RoboDK station: Estacion_Final_TFG.rdk

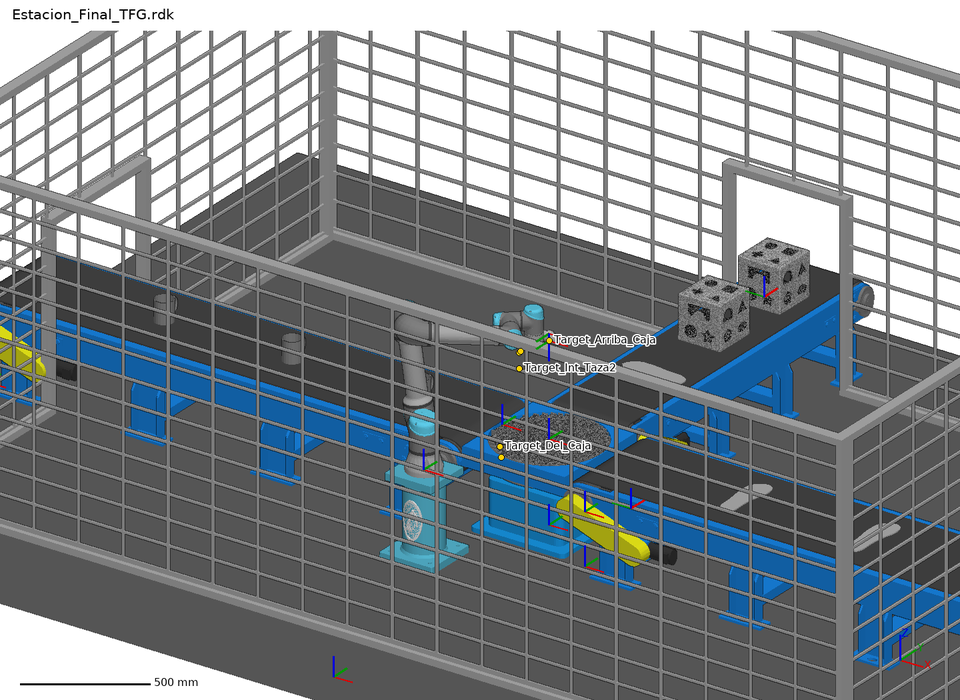
[picture v0: the station drawn from its stored meshes, robots at their saved joint values, targets as dots, program paths as lines]
Station Estacion_Final_TFG (saved by RoboDK 6.0.1). Poses are relative to the parent item; angles as X-Y-Z fixed-axis rotations.
Station parameters (name, value as stored): cara_actual, Cubo_Derecha, cam_delay, 0.005, contador, 10, prox_obj, Plantilla, defectuoso, 0, cont_def, 3, cont_ok, 4, prob_def, 5
  - folder Objetos
    - frame UR5e Base at (-167.75, -5.91, 0) mm
      - object Pedestal UR5 at (0, 0, -366.5) mm, size 250 x 250 x 366.5 mm, geometry from Pedestal-H12in-Type-1.sld
      - robot UR5e: 6 axes, payload 5 kg, reach 850 mm, repeatability 0.03 mm, weight 18.4 kg
          modified DH rows (alpha deg, a mm, theta deg, d mm): 0, 0, 0, 162.5; 90, 0, 180, 0; 0, 425, 0, 0; 0, 392.25, 0, 133.3; -90, 0, 0, 99.7; 90, 0, 180, 99.6
          joint limits [-360, -360, -360, -360, -360, -360] to [360, 360, 360, 360, 360, 360]; home [0, -90, -90, 0, 90, 0]; saved at [-138.346, -96.938, 101.969, -95.031, -90, -48.346]
        - frame Frame_Camara at (0, -105, 30.5) mm
          - camera Cámara 1
        - tool OnRobot Eyes Camera, TCP at (0.17, -105.19, 30.39) mm, size 104 x 155 x 41.9 mm
    - frame Frame_Cinta_Simple at (-2413.09, 275.71, -366.5) mm
      - robot Cinta_Simple: 1 axes
          modified DH rows (alpha deg, a mm, theta deg, d mm): 0, 0, 0, 0 linear
          base shift (0, 0, 0) mm, rotated rx 0 ry 90 rz 0 deg
          joint limits [-900000] to [900000]; home [0]; saved at [6082.39]
        - frame Frame_Padre_Cinta at (-2.39, 215, 0) mm
          - object Taza8 at (-4200, 0, 0) mm, rotated rx 0 ry 0 rz 90 deg, size 123.1 x 83.9 x 97 mm, geometry from Taza_Base.stp
          - object Taza9 at (-4800, 0, 0) mm, rotated rx 0 ry 0 rz 90 deg, size 123.1 x 83.9 x 97 mm, geometry from Taza_Base.stp
          - object Taza10 at (-5400, 0, 0) mm, rotated rx 0 ry 0 rz 90 deg, size 123.1 x 83.9 x 97 mm, geometry from Taza_Base.stp
    - frame Frame_Obj_Ref at (0, -850, -500) mm
      - object Juguete_ni at (0, 0, 0) mm, size 200 x 200 x 200 mm, geometry from Juguete_niños.stp
      - object Juguete_ni at (0, 0, 0) mm, size 200 x 200 x 200 mm, geometry from Juguete_niños_Arriba.stp
      - object Juguete_ni at (0, 0, 0) mm, size 200 x 200 x 200 mm, geometry from Juguete_niños_Der.stp
      - object Juguete_ni at (0, 0, 0) mm, size 200 x 200 x 200 mm, geometry from Juguete_niños_Frente.stp
      - object Juguete_ni at (0, 0, 0) mm, size 200 x 200 x 200 mm, geometry from Juguete_niños_Izq.stp
      - object Juguete_ni at (0, 0, 0) mm, size 200 x 200 x 200 mm, geometry from Juguete_niños_Det.stp
      - object Taza_Base at (0, 0, 0) mm, rotated rx 0 ry 0 rz 90 deg, size 123.1 x 83.9 x 97 mm, geometry from Taza_Base.stp
      - object Taza_Def1 at (0, 0, 0) mm, rotated rx 0 ry 0 rz 90 deg, size 123.1 x 83.9 x 97 mm, geometry from Taza_DibujoMal.stp
      - object Taza_Def2 at (0, 0, 0) mm, rotated rx 0 ry 0 rz 90 deg, size 123.1 x 83.9 x 97 mm, geometry from Taza_FaltaLetra.stp
      - object Plantilla_Derecha_Bien at (0, 0, 0) mm, rotated rx 90 ry 0 rz 0 deg, size 99.5 x 5 x 284.6 mm, geometry from Plantilla_Derecha_Bien.stl
      - object Plantilla_Derecha_Def1 at (0, 0, 0) mm, rotated rx 90 ry 0 rz 0 deg, size 99.6 x 5 x 284.5 mm, geometry from Plantilla_Derecha_Mal_Corte_Arriba.stl
      - object Plantilla_Derecha_Def2 at (0, 0, 0) mm, rotated rx 90 ry 0 rz 0 deg, size 99.6 x 5 x 284.6 mm, geometry from Plantilla_Derecha_Mal_Muescas.stl
      - object Plantilla_Izquierda_Bien at (0, 0, 0) mm, rotated rx 90 ry 0 rz 0 deg, size 99.5 x 5 x 284.6 mm, geometry from Plantilla_Izquierda_Bien.stl
      - object Plantilla_Izquierda_Def1 at (0, 0, 0) mm, rotated rx 90 ry 0 rz 0 deg, size 99.5 x 5 x 283.3 mm, geometry from Plantilla_Izquierda_Mal_Corte_Abajo.stl
      - object Plantilla_Izquierda_Def2 at (0, 0, 0) mm, rotated rx 90 ry 0 rz 0 deg, size 99.6 x 5 x 284.6 mm, geometry from Plantilla_Izquierda_Mal_Muescas.stl
    - frame Mesa_Rotatoria Base at (71.91, 490.71, -366.5) mm
      - robot Mesa_Rotatoria: 1 axes
          modified DH rows (alpha deg, a mm, theta deg, d mm): 0, 0, 0, 0
          joint limits [-360] to [360]; home [0]; saved at [0]
        - frame Cinta_Rotativa Base at (-220, 0, 366.5) mm
          - robot Cinta_Rotativa: 1 axes
              modified DH rows (alpha deg, a mm, theta deg, d mm): 0, 0, 0, 0 linear
              base shift (0, 0, 0) mm, rotated rx 0 ry 90 rz 0 deg
              joint limits [-10000] to [10000]; home [0]; saved at [3080]
      - object Base_Cinta at (0, 0, 280) mm, size 480 x 480 x 86.5 mm, geometry from Base_Cinta.stp
    - frame Frame_Cinta_OK at (391.91, 270.71, -366.5) mm
      - robot Cinta_OK: 1 axes
          modified DH rows (alpha deg, a mm, theta deg, d mm): 0, 0, 0, 0 linear
          base shift (0, 0, 0) mm, rotated rx 0 ry 90 rz 0 deg
          joint limits [-900000] to [900000]; home [0]; saved at [2400]
        - frame Frame_Padre_Cinta_OK at (-2.39, 215, 0) mm
          - object OK2 at (-600, 0, 0) mm, size 200 x 200 x 200 mm, geometry from Juguete_niños.stp
          - object OK3 at (-1200, 0, 0) mm, rotated rx 90 ry 0 rz 0 deg, size 99.5 x 5 x 284.6 mm, geometry from Plantilla_Izquierda_Bien.stl
          - object OK4 at (-1800, 0, 0) mm, rotated rx 90 ry 0 rz 0 deg, size 99.5 x 5 x 284.6 mm, geometry from Plantilla_Izquierda_Bien.stl
    - frame Frame_Cinta_Def at (247.91, 787.71, -366.5) mm, rotated rx 0 ry 0 rz 90 deg
      - robot Cinta_Def: 1 axes
          modified DH rows (alpha deg, a mm, theta deg, d mm): 0, 0, 0, 0 linear
          base shift (0, 0, 0) mm, rotated rx 0 ry 90 rz 0 deg
          joint limits [-900000] to [900000]; home [0]; saved at [1200]
        - frame Frame_Padre_Cinta_Def at (-2.39, 215, 0) mm
          - object Defectuoso1 at (0, -44, 0) mm, size 200 x 200 x 200 mm, geometry from Juguete_niños_Det.stp
          - object Defectuoso2 at (-400, -44, 0) mm, size 200 x 200 x 200 mm, geometry from Juguete_niños_Det.stp
          - object Defectuoso3 at (-800, -44, 0) mm, rotated rx 90 ry 0 rz 0 deg, size 99.6 x 5 x 284.5 mm, geometry from Plantilla_Derecha_Mal_Corte_Arriba.stl
    - frame Frame_Suelo at (117.25, 664.09, -367) mm
      - object Suelo at (0, 0, 0) mm, size 5420 x 3890 x 0 mm, geometry from Floor.sld
  - frame Frame_Targets at (71.91, 490.71, 450) mm, rotated rx 180 ry 0 rz 0 deg
    - target Target_Arriba_Caja (Cartesian target) at (0, 0, 30) mm; joints [-138.346, -96.938, 101.969, -95.031, -90, -48.346] of UR5e
    - target Target_Del_Caja (Cartesian target) at (0, 330, 350) mm, rotated rx 90 ry 0 rz 0 deg; joints [-204.685, -47.932, 150.066, -102.134, -24.685, -180] of UR5e
    - target Target_Int_Del (Cartesian target) at (0, 200, 0) mm; joints [-168.17, -117.089, 115.815, -88.726, -90, -78.17] of UR5e
    - target Target_Int_Taza1 (Cartesian target) at (0, 190, 0) mm; joints [-165.144, -119.371, 116.87, -87.498, -90, -75.144] of UR5e
    - target Target_Int_Taza2 (Cartesian target) at (0, 200, 70) mm, rotated rx 60 ry 0 rz 0 deg; joints [-180.443, -119.916, 146.516, -115.834, -30.003, -90.885] of UR5e
    - target Target_Taza (Cartesian target) at (0, 320, 400) mm, rotated rx 90 ry 0 rz 0 deg; joints [-202.098, -35.728, 146.743, -111.015, -22.098, -180] of UR5e
  - frame Frame_Target_Mesa at (71.91, 490.71, 0) mm
    - target Init_Mesa (Cartesian target) at (0, 0, 0) mm; joints [0, -47.932, 150.066, -102.134, -24.685, -180] of Mesa_Rotatoria
    - target Cubo_Izq (Cartesian target) at (0, 0, 0) mm, rotated rx 0 ry 0 rz 90 deg; joints [90, -47.932, 150.066, -102.134, -24.685, -180] of Mesa_Rotatoria
    - target Cubo_Detras (Cartesian target) at (0, 0, 0) mm, rotated rx 0 ry 0 rz 180 deg; joints [180, -47.932, 150.066, -102.134, -24.685, -180] of Mesa_Rotatoria
    - target Cubo_Der (Cartesian target) at (0, 0, 0) mm, rotated rx 0 ry 0 rz -90 deg; joints [270, -47.932, 150.066, -102.134, -24.685, -180] of Mesa_Rotatoria
    - target Target_Def (Cartesian target) at (0, 0, 0) mm, rotated rx 0 ry 0 rz 90 deg; joints [90, -47.932, 150.066, -102.134, -24.685, -180] of Mesa_Rotatoria
    - target Target_Taza_Mesa (Cartesian target) at (0, 0, 0) mm, rotated rx 0 ry 0 rz 90 deg; joints [90, -47.932, 150.066, -102.134, -24.685, -180] of Mesa_Rotatoria
  - folder Vallado
    - frame Frame Valla Trasera at (2332.25, -755.91, -366.5) mm, rotated rx 0 ry 0 rz 90 deg
      - object VallaTrasera at (0, 0, 0) mm, rotated rx 90 ry 0 rz 90 deg, size 4420 x 1500 x 50 mm, geometry from VallaBigCap.stl
    - frame Frame Valla Entrada at (-2062.75, -730.91, -366.5) mm, rotated rx 0 ry 0 rz -90 deg
      - object Valla_Entrada at (0, 0, 0) mm, rotated rx 90 ry 0 rz 180 deg, size 2790 x 1500 x 50 mm, geometry from Valla_Enrada.stp
    - frame Frame Valla Salida at (2307.25, -730.91, -366.5) mm, rotated rx 0 ry 0 rz -90 deg
      - object Valla_Salida at (0, 0, 0) mm, rotated rx 90 ry 0 rz 180 deg, size 2790 x 1500 x 50 mm, geometry from Valla_Enrada.stp
    - frame Frame Valla Defectuosas at (2332.25, 2084.09, -366.5) mm, rotated rx 0 ry 0 rz 180 deg
      - object Valla_CintaDef at (0, 0, 0) mm, rotated rx 90 ry 0 rz 0 deg, size 4420 x 1500 x 50 mm, geometry from Valla_CintaDef.stp
  - folder Programas
    - Python program Global (listed below)
    - Python program Reset (listed below)
  - folder Comparacion
    - Python program Comp_Inicial (listed below)
    - Python program Comp_Plantilla (listed below)
    - folder Codigos Cubo
      - Python program Comp_Cubo (listed below)
      - Python program Cubo_General (listed below)
    - folder Codigos Taza
      - Python program Comp_Taza (listed below)
      - Python program Taza_General (listed below)
  - folder Cintas
    - Python program Generar_Objeto (listed below)
    - Python program Avanzar_Cinta_Rot (listed below)

--- Python program Global ---
# Type help("robodk.robolink") or help("robodk.robomath") for more information
# Press F5 to run the script
# Documentation: https://robodk.com/doc/en/RoboDK-API.html
# Reference:     https://robodk.com/doc/en/PythonAPI/robodk.html
# Note: It is not required to keep a copy of this file, your Python script is saved with your RDK project

# You can also use the new version of the API:
from robodk import *      # RoboDK API
from robolink import *    # Robot toolbox
RDK = robolink.Robolink()

robot = RDK.Item('UR5e')
tool = RDK.Item('OnRobot Eyes Camera')
frame_target = RDK.Item('Frame_Targets')
init = RDK.Item('Reset')
avanzarCinta = RDK.Item('Generar_Objeto')
frame_mesa = RDK.Item('Frame_Target_Mesa')

arriba = RDK.Item('Target_Arriba_Caja')

robot.setPoseFrame(frame_target)
robot.MoveJ(arriba)

mesa=RDK.Item('Mesa_Rotatoria',itemtype=ITEM_TYPE_ROBOT)
cinta_rot=RDK.Item('Cinta_Rotativa',itemtype=ITEM_TYPE_ROBOT)
cinta_ok=RDK.Item('Cinta_OK',itemtype=ITEM_TYPE_ROBOT)
cinta_def=RDK.Item('Cinta_Def',itemtype=ITEM_TYPE_ROBOT)
ident = RDK.Item('Comp_Inicial')
comp_plantilla = RDK.Item('Comp_Plantilla')
comp_cubo = RDK.Item('Cubo_General')
comp_taza = RDK.Item('Taza_General')
avanzar_cinta_rot = RDK.Item('Avanzar_Cinta_Rot')
init_mesa = RDK.Item('Init_Mesa')
pos_def = RDK.Item('Target_Def')


frame_padre_def=RDK.Item('Frame_Padre_Cinta_Def')
frame_padre_ok=RDK.Item('Frame_Padre_Cinta_OK')

mesa.setPoseFrame(frame_mesa)

init.RunProgram()
init.WaitFinished()
obj_scan = RDK.getParam('prox_obj')

while True:
    while obj_scan == 'NULL':
        avanzarCinta.RunProgram()
        avanzarCinta.WaitFinished()
        obj_scan = RDK.getParam('prox_obj')

    avanzar_cinta_rot.RunProgram()
    avanzar_cinta_rot.WaitFinished()

    ident.RunProgram()
    ident.WaitFinished()

    defecto = RDK.getParam('defectuoso')
    contador = int(RDK.getParam('contador'))
    contador_def = int(RDK.getParam('cont_def'))
    contador_ok = int(RDK.getParam('cont_ok'))
    nombre_obj = obj_scan+str(contador-3)
    obj_listo = RDK.Item(nombre_obj)

    if defecto == 1:
        mesa.MoveJ(pos_def)
        avanzar_cinta_rot.RunProgram()
        avanzar_cinta_rot.WaitFinished()
        obj_listo.setParent(frame_padre_def)
        if obj_scan == 'Plantilla':
            obj_listo.setPose(transl((-400*(contador_def)),-44,0) * rotx(pi/2))
        elif obj_scan == 'Taza':
            obj_listo.setPose(transl((-400*(contador_def)),-44,0) * rotz(pi/2))
        else:
            obj_listo.setPose(transl((-400*(contador_def)),-44,0))
        cinta_def.MoveJ(cinta_def.Joints()+400)
        contador_def += 1
        obj_listo.setName('Defectuoso'+str(contador_def))
        if contador_def > 3:
            obj_borrar = RDK.Item('Defectuoso'+str(contador_def-3))
            RDK.Delete(obj_borrar)

    else:
        mesa.MoveJ(init_mesa)
        avanzar_cinta_rot.RunProgram()
        avanzar_cinta_rot.WaitFinished()
        obj_listo.setParent(frame_padre_ok)
        if obj_scan == 'Plantilla':
            obj_listo.setPose(transl((-600*(contador_ok)),0,0) * rotx(pi/2))
        elif obj_scan == 'Taza':
            obj_listo.setPose(transl((-600*(contador_ok)),0,0) * rotz(pi/2))
        else:
            obj_listo.setPose(transl((-600*(contador_ok)),0,0))
        cinta_ok.MoveJ(cinta_ok.Joints()+600)
        contador_ok += 1
        obj_listo.setName('OK'+str(contador_ok))
        if contador_ok > 3:
            obj_borrar = RDK.Item('OK'+str(contador_ok-3))
            RDK.Delete(obj_borrar)

    RDK.setParam('cont_def',contador_def)
    RDK.setParam('cont_ok',contador_ok)
    mesa.MoveJ(init_mesa)
    RDK.setParam('defectuoso',0)
    avanzarCinta.RunProgram()
    avanzarCinta.WaitFinished()
    obj_scan = RDK.getParam('prox_obj')

--- Python program Reset ---
# Type help("robodk.robolink") or help("robodk.robomath") for more information
# Press F5 to run the script
# Documentation: https://robodk.com/doc/en/RoboDK-API.html
# Reference:     https://robodk.com/doc/en/PythonAPI/robodk.html
# Note: It is not required to keep a copy of this file, your Python script is saved with your RDK project

import random

# Forward and backwards compatible use of the RoboDK API:
# Remove these 2 lines to follow python programming guidelines
from robodk import *      # RoboDK API
from robolink import *    # Robot toolbox
# Link to RoboDK
RDK = Robolink()

num=random.randint(1,3)
#num=3

RDK.setParam('contador',1)
RDK.setParam('cont_def',0)
RDK.setParam('cont_ok',0)
RDK.setParam('defectuoso',0)

if num == 1: # Caso de que sea plantilla
    num2 = random.randint(1,2)
    if num2 == 1: # Plantilla izquierda
        num3 = random.randint(1,6)
        if num3 == 5: # Defecto 1
            padre = RDK.Item('Plantilla_Izquierda_Def1')
            nombreCopia = 'Plantilla'
        elif num3 == 6: # Defecto 2
            padre = RDK.Item('Plantilla_Izquierda_Def2')
            nombreCopia = 'Plantilla'
        else:
            padre = RDK.Item('Plantilla_Izquierda_Bien')
            nombreCopia = 'Plantilla'
    if num2 == 2: # Plantilla izquierda
        num3 = random.randint(1,6)
        if num3 == 5: # Defecto 1
            padre = RDK.Item('Plantilla_Derecha_Def1')
            nombreCopia = 'Plantilla'
        elif num3 == 6: # Defecto 2
            padre = RDK.Item('Plantilla_Derecha_Def2')
            nombreCopia = 'Plantilla'
        else:
            padre = RDK.Item('Plantilla_Derecha_Bien')
            nombreCopia = 'Plantilla'

elif num == 2: # Caso de que sea Juguete
    num2 = random.randint(1,10)
    if num2 == 6: # Juguete mal arriba
        padre = RDK.Item('Juguete_niños_Arriba')
        nombreCopia = 'Juguete_niños'
    elif num2 == 7: # Juguete mal izquierda
        padre = RDK.Item('Juguete_niños_Izq')
        nombreCopia = 'Juguete_niños'
    elif num2 == 8: # Juguete mal derecha
        padre = RDK.Item('Juguete_niños_Der')
        nombreCopia = 'Juguete_niños'
    elif num2 == 9: # Juguete mal delante
        padre = RDK.Item('Juguete_niños_Del')
        nombreCopia = 'Juguete_niños'
    elif num2 == 10: # Juguete mal detras
        padre = RDK.Item('Juguete_niños_Det')
        nombreCopia = 'Juguete_niños'
    else: # Caso sin fallos
        padre = RDK.Item('Juguete_niños_Base')
        nombreCopia = 'Juguete_niños'

elif num == 3: # Caso de que sea taza
    num2 = random.randint(1,6)
    if num2 == 5: # Defecto 1
        padre = RDK.Item('Taza_Def1')
        nombreCopia = 'Taza'
    elif num2 == 6: # Defecto 2
        padre = RDK.Item('Taza_Def2')
        nombreCopia = 'Taza'
    else:
        padre = RDK.Item('Taza_Base')
        nombreCopia = 'Taza'


MECHANISM_NAME = 'Cinta_Simple'
mechanism=RDK.Item(MECHANISM_NAME,itemtype=ITEM_TYPE_ROBOT)
cinta_ok=RDK.Item('Cinta_OK',itemtype=ITEM_TYPE_ROBOT)
cinta_def=RDK.Item('Cinta_Def',itemtype=ITEM_TYPE_ROBOT)
cinta_rot=RDK.Item('Cinta_Rotativa',itemtype=ITEM_TYPE_ROBOT)
frame_padre_def=RDK.Item('Frame_Padre_Cinta_Def')
frame_padre_ok=RDK.Item('Frame_Padre_Cinta_OK')
mesa = RDK.Item('Mesa_Rotatoria')

frame_padre=RDK.Item('Frame_Padre_Cinta')

if mechanism.Valid() and cinta_rot.Valid() and mesa.Valid():
    mechanism.setJoints([467.39])
    cinta_ok.setJoints([0])
    cinta_def.setJoints([0])
    cinta_rot.setJoints([0])
    mesa.setJoints([0])
    RDK.Delete(frame_padre.Childs())
    RDK.Delete(frame_padre_def.Childs())
    RDK.Delete(frame_padre_ok.Childs())
    RDK.Delete(cinta_rot.Childs())
    padre.Copy()
    copia=RDK.Paste()
    copia.setParent(frame_padre)
    RDK.setParam('prox_obj','NULL')
    #hacemos visible el objeto nuevo
    cont = int(RDK.getParam('contador'))
    copia.setName(nombreCopia+str(cont))
    copia.setVisible(1)

--- Python program Comp_Inicial ---
from robolink import *
import cv2 as cv
import numpy as np
import os

RDK = Robolink()
cam_item = RDK.Item('Cámara 1', ITEM_TYPE_CAMERA)
carpeta = r"C:\Users\algob\OneDrive\UPV\4 - Cuarto\TFG\Imagen"

comp_plantilla = RDK.Item('Comp_Plantilla')
comp_cubo = RDK.Item('Cubo_General')
comp_taza = RDK.Item('Taza_General')

# 1. Cargar las dos imagenes de referencia en escala de grises (RAW)
img_izq_raw = cv.imread(os.path.join(carpeta, "Ref_izq.png"), 0)
img_der_raw = cv.imread(os.path.join(carpeta, "Ref_der.png"), 0)
img_cubo_raw = cv.imread(os.path.join(carpeta, "Cubo", "Cubo_Arriba_base.png"), 0)
img_taza_raw = cv.imread(os.path.join(carpeta, "Taza", "Taza_Arriba.png"), 0)

# FILTRO: Convertir el fondo gris en NEGRO puro y la plantilla en BLANCO puro
_, img_izq = cv.threshold(img_izq_raw, 200, 255, cv.THRESH_BINARY)
_, img_der = cv.threshold(img_der_raw, 200, 255, cv.THRESH_BINARY)
_, img_cubo = cv.threshold(img_cubo_raw, 200, 255, cv.THRESH_BINARY)
_, img_taza = cv.threshold(img_taza_raw, 200, 255, cv.THRESH_BINARY)

def obtener_contorno_principal(img_bw):
    # RETR_EXTERNAL busca únicamente el contorno exterior más externo
    cnts, _ = cv.findContours(img_bw, cv.RETR_EXTERNAL, cv.CHAIN_APPROX_SIMPLE)
    return max(cnts, key=cv.contourArea) if cnts else None

ref_izq = obtener_contorno_principal(img_izq)
ref_der = obtener_contorno_principal(img_der)
ref_cubo = obtener_contorno_principal(img_cubo)
ref_taza = obtener_contorno_principal(img_taza)

tiempo_inicio = time.time()
DURACION_MAXIMA = RDK.getParam('cam_delay')

while True:
    if (time.time() - tiempo_inicio) > DURACION_MAXIMA:
        cv.destroyAllWindows()
        cv.waitKey(1)
        break

    bytes_img = RDK.Cam2D_Snapshot("", cam_item)
    if bytes_img == b'':
        cv.destroyAllWindows()
        cv.waitKey(1)
        break

    img = cv.imdecode(np.frombuffer(bytes_img, np.uint8), cv.IMREAD_UNCHANGED)
    gray = cv.cvtColor(img, cv.COLOR_BGR2GRAY)

    _, thresh = cv.threshold(gray, 200, 255, cv.THRESH_BINARY)
    actual = obtener_contorno_principal(thresh)

    if actual is not None:
        diff_izq = cv.matchShapes(ref_izq, actual, 1, 0.0)
        diff_der = cv.matchShapes(ref_der, actual, 1, 0.0)
        diff_cubo = cv.matchShapes(ref_cubo, actual, 1, 0.0)
        diff_taza = cv.matchShapes(ref_taza, actual, 1, 0.0)

        mejor_diff = min(diff_izq, diff_der, diff_taza, diff_cubo)

        if mejor_diff == diff_izq or mejor_diff == diff_der:
            comp_plantilla.RunProgram()
            comp_plantilla.WaitFinished()
        elif mejor_diff == diff_cubo:
            comp_cubo.RunProgram()
            comp_cubo.WaitFinished()
        elif mejor_diff == diff_taza:
            comp_taza.RunProgram()
            comp_taza.WaitFinished()

cv.destroyAllWindows()
cv.waitKey(1)

--- Python program Comp_Plantilla ---
from robolink import *
import cv2 as cv
import numpy as np
import os

RDK = Robolink()
cam_item = RDK.Item('Cámara 1', ITEM_TYPE_CAMERA)
carpeta = r"C:\Users\algob\OneDrive\UPV\4 - Cuarto\TFG\Imagen"

# 1. Cargar las dos imagenes de referencia en escala de grises (RAW)
img_izq_raw = cv.imread(os.path.join(carpeta, "Ref_izq.png"), 0)
img_der_raw = cv.imread(os.path.join(carpeta, "Ref_der.png"), 0)

# FILTRO: Convertir el fondo gris en NEGRO puro y la plantilla en BLANCO puro
_, img_izq = cv.threshold(img_izq_raw, 200, 255, cv.THRESH_BINARY)
_, img_der = cv.threshold(img_der_raw, 200, 255, cv.THRESH_BINARY)

def obtener_contorno_principal(img_bw):
    # RETR_EXTERNAL busca únicamente el contorno exterior más externo
    cnts, _ = cv.findContours(img_bw, cv.RETR_EXTERNAL, cv.CHAIN_APPROX_SIMPLE)
    return max(cnts, key=cv.contourArea) if cnts else None

ref_izq = obtener_contorno_principal(img_izq)
ref_der = obtener_contorno_principal(img_der)

# Umbral de aceptación
UMBRAL = 0.01
tiempo_inicio = time.time()
DURACION_MAXIMA = RDK.getParam('cam_delay')

while True:
    if (time.time() - tiempo_inicio) > DURACION_MAXIMA:
        cv.destroyAllWindows()
        cv.waitKey(1)
        break

    bytes_img = RDK.Cam2D_Snapshot("", cam_item)
    if bytes_img == b'':
        cv.destroyAllWindows()
        cv.waitKey(1)
        break

    img = cv.imdecode(np.frombuffer(bytes_img, np.uint8), cv.IMREAD_UNCHANGED)
    gray = cv.cvtColor(img, cv.COLOR_BGR2GRAY)

    _, thresh = cv.threshold(gray, 200, 255, cv.THRESH_BINARY)
    actual = obtener_contorno_principal(thresh)

    if actual is not None:
        # 2. Comparar con ambas imagenes de referencia
        diff_izq = cv.matchShapes(ref_izq, actual, 1, 0.0)
        diff_der = cv.matchShapes(ref_der, actual, 1, 0.0)

        # Elegir la que mejor encaje (menor valor)
        mejor_diff = min(diff_izq, diff_der)

        # Seleccionar la imagen de fondo de referencia correcta según la forma detectada
        if diff_izq < diff_der:
            img_ref_base = img_izq.copy()
            contorno_ref = ref_izq
        else:
            img_ref_base = img_der.copy()
            contorno_ref = ref_der

        # Crear la ventana de la Imagen de Referencia
        # Convertimos la referencia a BGR para poder dibujarle la línea en color azul
        img_referencia_color = cv.cvtColor(img_ref_base, cv.COLOR_GRAY2BGR)
        cv.drawContours(img_referencia_color, [contorno_ref], -1, (255, 0, 0), 2)
        cv.imshow("Ref", img_referencia_color)

        # 3. Lógica de decisión para la pieza actual
        if mejor_diff < UMBRAL:
            color, estado = (0, 255, 0), "OK -"
        else:
            color, estado = (0, 0, 255), "DEFECTUOSA -"
            RDK.setParam('defectuoso',1)

        # Dibujar contorno verde/rojo en la imagen de la cámara
        cv.drawContours(img, [actual], -1, color, 2)
        cv.putText(img, f"{estado} ({mejor_diff:.3f})", (5, 40),
                    cv.FONT_HERSHEY_SIMPLEX, 0.7, color, 2)

    cv.imshow("Inspección", img)

    key = cv.waitKey(30) & 0xFF
    if key == 27: # Tecla ESC para salir
        break

    # Control de cierre si el usuario cierra cualquiera de las dos ventanas con la 'X'
    if (cv.getWindowProperty("Inspección", cv.WND_PROP_VISIBLE) < 1 or
        cv.getWindowProperty("Ref", cv.WND_PROP_VISIBLE) < 1):
        break

cv.destroyAllWindows()
cv.waitKey(1)

--- Python program Comp_Cubo ---
from robolink import *
import cv2 as cv
import numpy as np
import os
import time

RDK = Robolink()
cam_item = RDK.Item('Cámara 1', ITEM_TYPE_CAMERA)
carpeta_base = r"C:\Users\algob\OneDrive\UPV\4 - Cuarto\TFG\Imagen\Cubo"

# 1. CARGAR Y PROCESAR LA IMAGEN ref DE REFERENCIA
nombre_ref = RDK.getParam("cara_actual") + "_base.png"
ruta_ref = os.path.join(carpeta_base, nombre_ref)
img_ref_raw = cv.imread(ruta_ref, 0)

def obtener_contornos_internos(img_bw):
    cnts, _ = cv.findContours(img_bw, cv.RETR_LIST, cv.CHAIN_APPROX_SIMPLE)

    figuras_internas = []
    for c in cnts:
        area = cv.contourArea(c)
        if 4000 < area < 40000:
            figuras_internas.append(c)

    return figuras_internas

def calcular_hu_global(img_bw, contornos):
    mascara = np.zeros_like(img_bw)
    cv.drawContours(mascara, contornos, -1, 255, -1)
    momentos = cv.moments(mascara)
    hu = cv.HuMoments(momentos).flatten()
    hu_log = -np.sign(hu) * np.log10(np.abs(hu))
    return hu_log



if img_ref_raw is None:
    RDK.ShowMessage(f"ERROR: No se encontró la imagen de referencia en: {ruta_ref}")
else:
    _, thresh_ref = cv.threshold(img_ref_raw, 100, 255, cv.THRESH_BINARY_INV)

    if np.sum(thresh_ref[0:10, 0:10]) > 200000:
        _, thresh_ref = cv.threshold(img_ref_raw, 100, 255, cv.THRESH_BINARY)

    cnts_ref = obtener_contornos_internos(thresh_ref)
    hu_ref = calcular_hu_global(thresh_ref, cnts_ref)

# Umbral de tolerancia
UMBRAL = 0.3

# --- CONTROL DE TIEMPO PRINCIPAL ---
tiempo_inicio = time.time()
DURACION_MAXIMA = RDK.getParam('cam_delay')

while True:
    if (time.time() - tiempo_inicio) > DURACION_MAXIMA:
        cv.destroyAllWindows()
        cv.waitKey(1)
        break

    bytes_img = RDK.Cam2D_Snapshot("", cam_item)
    if bytes_img == b'':
        cv.destroyAllWindows()
        cv.waitKey(1)
        break

    img = cv.imdecode(np.frombuffer(bytes_img, np.uint8), cv.IMREAD_UNCHANGED)
    gray = cv.cvtColor(img, cv.COLOR_BGR2GRAY)

    _, thresh_actual = cv.threshold(gray, 100, 255, cv.THRESH_BINARY_INV)
    if np.sum(thresh_actual[0:10, 0:10]) > 200000:
        _, thresh_actual = cv.threshold(gray, 100, 255, cv.THRESH_BINARY)

    if img_ref_raw is not None:
        cnts_actuales = obtener_contornos_internos(thresh_actual)

        if len(cnts_actuales) > 0:
            hu_actual = calcular_hu_global(thresh_actual, cnts_actuales)
            dif = np.linalg.norm(hu_ref - hu_actual)

            if dif < UMBRAL:
                color, estado_texto = (0, 255, 0), "CARA OK -"
            else:
                color, estado_texto = (0, 0, 255), "DEFECTO -"
                RDK.setParam("defectuoso",1)

            # DIBUJAMOS EL BORDE DIRECTAMENTE EN LAS FORMAS INTERIORES
            cv.drawContours(img, cnts_actuales, -1, color, 2)
            cv.putText(img, f"{estado_texto} (Diff: {dif:.4f})", (15, 40),
                        cv.FONT_HERSHEY_SIMPLEX, 0.6, color, 2)
        else:
            cv.putText(img, "PATRONES NO DETECTADOS", (15, 40),
                        cv.FONT_HERSHEY_SIMPLEX, 0.6, (255, 165, 0), 2)

        # Ventana Secundaria: Mostrar ref con sus patrones marcados en AZUL
        img_ref_visual = cv.cvtColor(thresh_ref, cv.COLOR_GRAY2BGR)
        if 'cnts_ref' in locals():
            cv.drawContours(img_ref_visual, cnts_ref, -1, (255, 0, 0), 2)
        cv.imshow("Ref", img_ref_visual)

    cv.imshow("Inspeccion", img)

    # El waitKey es vital para refrescar la interfaz gráfica de OpenCV
    key = cv.waitKey(30) & 0xFF
    if key == 27: # ESC
        cv.destroyAllWindows()
        cv.waitKey(1)
        break

    if (cv.getWindowProperty("Inspeccion", cv.WND_PROP_VISIBLE) < 1 or
        cv.getWindowProperty("Ref", cv.WND_PROP_VISIBLE) < 1):
        cv.destroyAllWindows()
        cv.waitKey(1)
        break

# Cierre final de seguridad y reporte a RoboDK
cv.destroyAllWindows()
cv.waitKey(1)

--- Python program Cubo_General ---
# Forward and backwards compatible use of the RoboDK API:
# Remove these 2 lines to follow python programming guidelines
from robodk import *      # RoboDK API
from robolink import *    # Robot toolbox
# Link to RoboDK

RDK = Robolink()
robot = RDK.Item('UR5e')
mesa = RDK.Item('Mesa_Rotatoria')
frame_target = RDK.Item('Frame_Targets')
frame_mesa = RDK.Item('Frame_Target_Mesa')
tool = RDK.Item('OnRobot Eyes Camera')

arriba = RDK.Item('Target_Arriba_Caja')
int_del = RDK.Item('Target_Int_Del')
delante = RDK.Item('Target_Del_Caja')

cubo_izq = RDK.Item('Cubo_Izq')
cubo_der = RDK.Item('Cubo_Der')
cubo_det = RDK.Item('Cubo_Detras')
init_mesa = RDK.Item('Init_Mesa')

#avanzar = RDK.Item('Avanzar_Cinta')
inspeccion = RDK.Item('Comp_Cubo')

actual = RDK.getParam('cara_actual')

robot.setPoseFrame(frame_target)
mesa.setPoseFrame(frame_mesa)

robot.MoveJ(arriba)
RDK.setParam('cara_actual','Cubo_Arriba')
inspeccion.RunProgram()
inspeccion.WaitFinished()

fallo = RDK.getParam("defectuoso")
if fallo == 0:
    robot.MoveL(int_del)
    robot.MoveJ(delante)
    RDK.setParam('cara_actual','Cubo_Delante')
    inspeccion.RunProgram()
    inspeccion.WaitFinished()

    fallo = RDK.getParam("defectuoso")
    if fallo == 0:
        mesa.MoveJ(cubo_izq)
        RDK.setParam('cara_actual','Cubo_Izquierda')
        inspeccion.RunProgram()
        inspeccion.WaitFinished()


        fallo = RDK.getParam("defectuoso")
        if fallo == 0:
            mesa.MoveJ(cubo_det)
            RDK.setParam('cara_actual','Cubo_Detras')
            inspeccion.RunProgram()
            inspeccion.WaitFinished()

            fallo = RDK.getParam("defectuoso")
            if fallo == 0:
                mesa.MoveJ(cubo_der)
                RDK.setParam('cara_actual','Cubo_Derecha')
                inspeccion.RunProgram()
                inspeccion.WaitFinished()
                robot.MoveJ(int_del)
                fallo = RDK.getParam("defectuoso")
                if fallo == 0:
                    mesa.MoveJ(init_mesa)
            else:
                robot.MoveJ(int_del)
        else:
            robot.MoveJ(int_del)
    else:
        robot.MoveJ(int_del)

robot.MoveL(arriba)

--- Python program Comp_Taza ---
from robodk import robolink    # RoboDK API
from robodk import robomath    # Robot toolbox
import cv2 as cv
import numpy as np
import os
import time
from robolink import *

RDK = Robolink()
cam_item = RDK.Item('Cámara 1', ITEM_TYPE_CAMERA)
carpeta_base = r"C:\Users\algob\OneDrive\UPV\4 - Cuarto\TFG\Imagen\Taza"

# 1. CARGAR Y PROCESAR LA IMAGEN DE REFERENCIA DE LA TAZA
img_ref_raw = cv.imread(os.path.join(carpeta_base, "Taza_Base.png"), 0)

def obtener_contornos_logo(img_bw):
    # RETR_TREE devuelve la jerarquía completa [Next, Previous, Child, Parent]
    cnts, hierarchy = cv.findContours(img_bw, cv.RETR_TREE, cv.CHAIN_APPROX_SIMPLE)

    figuras_logo = []
    if hierarchy is None:
        return figuras_logo

    hierarchy = hierarchy[0]

    for i, c in enumerate(cnts):
        area = cv.contourArea(c)
        if 60 < area < 30000:
            padre_idx = hierarchy[i][3]
            if padre_idx != -1:
                x, y, w, h = cv.boundingRect(c)
                proporcion = w / float(h)
                if proporcion < 3.0:
                    figuras_logo.append(c)

    return figuras_logo

def calcular_hu_global(img_bw, contornos):
    mascara = np.zeros_like(img_bw)
    cv.drawContours(mascara, contornos, -1, 255, -1)
    momentos = cv.moments(mascara)
    hu = cv.HuMoments(momentos).flatten()
    hu_log = -np.sign(hu) * np.log10(np.abs(hu))
    return hu_log


if img_ref_raw is None:
    RDK.ShowMessage(f"ERROR: No se encontró la imagen de referencia en: {carpeta_base}")
else:
    _, thresh_ref = cv.threshold(img_ref_raw, 60, 255, cv.THRESH_BINARY)

    if np.sum(thresh_ref[0:10, 0:10]) > 200000:
        _, thresh_ref = cv.threshold(img_ref_raw, 60, 255, cv.THRESH_BINARY_INV)

    cnts_ref = obtener_contornos_logo(thresh_ref)
    hu_ref = calcular_hu_global(thresh_ref, cnts_ref)

# Umbral de tolerancia para la verificación del Logotipo
UMBRAL = 0.1

# --- CONTROL DE TIEMPO PRINCIPAL (5 SEGUNDOS) ---
tiempo_inicio = time.time()
DURACION_MAXIMA = RDK.getParam('cam_delay')

ultimo_estado = "SIN DETECCIÓN"

while True:
    if (time.time() - tiempo_inicio) > DURACION_MAXIMA:
        cv.destroyAllWindows()
        cv.waitKey(1)
        break

    bytes_img = RDK.Cam2D_Snapshot("", cam_item)
    if bytes_img == b'':
        cv.destroyAllWindows()
        cv.waitKey(1)
        break

    img = cv.imdecode(np.frombuffer(bytes_img, np.uint8), cv.IMREAD_UNCHANGED)
    gray = cv.cvtColor(img, cv.COLOR_BGR2GRAY)

    # Binarización de la imagen
    _, thresh_actual = cv.threshold(gray, 60, 255, cv.THRESH_BINARY)
    # Si hay muchos píxeles blancos se hace una binarización invertida
    if np.sum(thresh_actual[0:10, 0:10]) > 200000:
        _, thresh_actual = cv.threshold(gray, 60, 255, cv.THRESH_BINARY_INV)

    if img_ref_raw is not None:
        cnts_actuales = obtener_contornos_logo(thresh_actual)

        if len(cnts_actuales) > 0:
            hu_actual = calcular_hu_global(thresh_actual, cnts_actuales)
            dif = np.linalg.norm(hu_ref - hu_actual)

            if dif < UMBRAL:
                color, estado_texto = (0, 255, 0), "LOGO OK -"
                ultimo_estado = f"CORRECTA (Diff: {dif:.4f})"
            else:
                color, estado_texto = (0, 0, 255), "DEFECTO -"
                ultimo_estado = f"DEFECTO (Diff: {dif:.4f})"
                RDK.setParam("defectuoso", 1)

            # Pintar los componentes del logotipo en verde/rojo
            cv.drawContours(img, cnts_actuales, -1, color, 2)
            cv.putText(img, f"{estado_texto} (Diff: {dif:.4f})", (15, 40),
                        cv.FONT_HERSHEY_SIMPLEX, 0.6, color, 2)
        else:
            ultimo_estado = "LOGO NO DETECTADO"
            cv.putText(img, "BUSCANDO LOGO...", (15, 40),
                        cv.FONT_HERSHEY_SIMPLEX, 0.6, (255, 165, 0), 2)

        # Ventana de Referencia del modelo maestro de la taza
        img_ref_visual = cv.cvtColor(thresh_ref, cv.COLOR_GRAY2BGR)
        if 'cnts_ref' in locals():
            cv.drawContours(img_ref_visual, cnts_ref, -1, (255, 0, 0), 2)

        cv.imshow("Ref", img_ref_visual)

    cv.imshow("Inspección", img)

    key = cv.waitKey(30) & 0xFF
    if key == 27:
        cv.destroyAllWindows()
        cv.waitKey(1)
        break

    if (cv.getWindowProperty("Inspección", cv.WND_PROP_VISIBLE) < 1 or
        cv.getWindowProperty("Ref", cv.WND_PROP_VISIBLE) < 1):
        cv.destroyAllWindows()
        cv.waitKey(1)
        break

# Cierre ordenado y reporte a la terminal de RoboDK
cv.destroyAllWindows()
cv.waitKey(1)

--- Python program Taza_General ---
# Forward and backwards compatible use of the RoboDK API:
# Remove these 2 lines to follow python programming guidelines
from robodk import *      # RoboDK API
from robolink import *    # Robot toolbox
# Link to RoboDK

RDK = Robolink()
robot = RDK.Item('UR5e')
mesa = RDK.Item('Mesa_Rotatoria')
frame_target = RDK.Item('Frame_Targets_Taza')
frame_base = RDK.Item('Frame_Targets')
frame_mesa = RDK.Item('Frame_Target_Mesa')
tool = RDK.Item('OnRobot Eyes Camera')
cinta = RDK.Item('Cinta_Rotativa',itemtype=ITEM_TYPE_ROBOT)

arriba = RDK.Item('Target_Arriba_Caja')
int_1 = RDK.Item('Target_Int_Taza1')
int_2 = RDK.Item('Target_Int_Taza2')
taza = RDK.Item('Target_Taza')

taza_mesa = RDK.Item('Target_Taza_Mesa')
init_mesa = RDK.Item('Init_Mesa')

inspeccion = RDK.Item('Comp_Taza')


robot.setPoseFrame(frame_target)
mesa.setPoseFrame(frame_mesa)

robot.MoveL(int_1)
robot.MoveJ(int_2)
robot.MoveJ(taza)
mesa.MoveJ(taza_mesa)
cinta.MoveJ(cinta.Joints()-180)
inspeccion.RunProgram()
inspeccion.WaitFinished()
cinta.MoveJ(cinta.Joints()+180)
robot.MoveJ(int_2)
robot.MoveJ(int_1)
robot.setPoseFrame(frame_base)
robot.MoveL(arriba)

--- Python program Generar_Objeto ---
import random
from robodk import *      # RoboDK API
from robolink import *    # Robot toolbox

RDK = Robolink()

MECHANISM_NAME='Cinta_Simple'
INCREMENTO_MM=600

#Obtenemos el valor de la variable contador la cual está definida en la estación
contador=int(RDK.getParam('contador'))
mechanism=RDK.Item(MECHANISM_NAME,itemtype=ITEM_TYPE_ROBOT)
cinta_rot=RDK.Item('Cinta_Rotativa',itemtype=ITEM_TYPE_ROBOT)

num = random.randint(1,3)
#num = 3 # Debug para generar solo un tipo de objeto

if num == 1: # Caso de que sea plantilla
    num2 = random.randint(1,2)
    if num2 == 1: # Plantilla izquierda
        num3 = random.randint(1,6)
        if num3 == 5: # Defecto 1
            padre = RDK.Item('Plantilla_Izquierda_Def1')
            nombreCopia = 'Plantilla'
        elif num3 == 6: # Defecto 2
            padre = RDK.Item('Plantilla_Izquierda_Def2')
            nombreCopia = 'Plantilla'
        else:
            padre = RDK.Item('Plantilla_Izquierda_Bien')
            nombreCopia = 'Plantilla'
    if num2 == 2: # Plantilla izquierda
        num3 = random.randint(1,6)
        if num3 == 5: # Defecto 1
            padre = RDK.Item('Plantilla_Derecha_Def1')
            nombreCopia = 'Plantilla'
        elif num3 == 6: # Defecto 2
            padre = RDK.Item('Plantilla_Derecha_Def2')
            nombreCopia = 'Plantilla'
        else:
            padre = RDK.Item('Plantilla_Derecha_Bien')
            nombreCopia = 'Plantilla'

elif num == 2: # Caso de que sea Juguete
    num2 = random.randint(1,10) # Modo normal
    #num2 = random.randint(6,10) # Modo solo defectuosos
    if num2 == 6: # Juguete mal arriba
        padre = RDK.Item('Juguete_niños_Arriba')
        nombreCopia = 'Juguete_niños'
    elif num2 == 7: # Juguete mal izquierda
        padre = RDK.Item('Juguete_niños_Izq')
        nombreCopia = 'Juguete_niños'
    elif num2 == 8: # Juguete mal derecha
        padre = RDK.Item('Juguete_niños_Der')
        nombreCopia = 'Juguete_niños'
    elif num2 == 9: # Juguete mal delante
        padre = RDK.Item('Juguete_niños_Del')
        nombreCopia = 'Juguete_niños'
    elif num2 == 10: # Juguete mal detras
        padre = RDK.Item('Juguete_niños_Det')
        nombreCopia = 'Juguete_niños'
    else: # Caso sin fallos
        padre = RDK.Item('Juguete_niños_Base')
        nombreCopia = 'Juguete_niños'

elif num == 3: # Caso de que sea taza
    num2 = random.randint(1,6)
    if num2 == 5: # Defecto 1
        padre = RDK.Item('Taza_Def1')
        nombreCopia = 'Taza'
    elif num2 == 6: # Defecto 2
        padre = RDK.Item('Taza_Def2')
        nombreCopia = 'Taza'
    else:
        padre = RDK.Item('Taza_Base')
        nombreCopia = 'Taza'


#Este es el sistema de referencia en el que meteremos el elemento copiado
frame_padre=RDK.Item('Frame_Padre_Cinta')

plantilla = RDK.Item('Plantilla' + str(int(contador - 2)))
juguete = RDK.Item('Juguete_niños' + str(int(contador - 2)))
taza = RDK.Item('Taza' + str(int(contador - 2)))

if mechanism.Valid():

    #Avanzamos la cinta
    mechanism.MoveJ(mechanism.Joints()+INCREMENTO_MM)
    #Copiamos el objeto
    padre.Copy()
    #Pegamos el objeto
    copia=RDK.Paste()
    #Lo metemos en el sistema de referencia donde estarán todos los objetos
    copia.setParent(frame_padre)
    #incrementamos la cuenta de objetos copiados
    contador=contador+1
    #Cambiamos la posición del elemento copiado haciendo una traslación que corresponde
    #en el eje X a el número de veces que hemos hecho avanzar ya la cinta
    if num == 1: # si se genera una plantilla
        copia.setPose(transl((-INCREMENTO_MM)*(contador-1),0,0) * rotx(pi/2))
    elif num == 3:
        copia.setPose(transl((-INCREMENTO_MM)*(contador-1),0,0) * rotz(pi/2))
    else:
        copia.setPose(transl((-INCREMENTO_MM)*(contador-1),0,0))

    #hacemos visible el objeto nuevo
    copia.setName(nombreCopia + str(int(contador)))
    copia.setVisible(1)
    #Actualizamos el valor de la variable contador en la estación
    RDK.setParam('contador',contador)

    #Determinamos que objeto va a llegar a la cinta rotatoria
    if plantilla.Valid():
        RDK.setParam('prox_obj','Plantilla')
        plantilla.setParent(cinta_rot)
        plantilla.setPose(transl((-440*(contador-4)),0,0) * rotx(pi/2))


    elif juguete.Valid():
        RDK.setParam('prox_obj','Juguete_niños')
        juguete.setParent(cinta_rot)
        juguete.setPose(transl((-440*(contador-4)),0,0))

    elif taza.Valid():
        RDK.setParam('prox_obj','Taza')
        taza.setParent(cinta_rot)
        taza.setPose(transl((-440*(contador-4)),0,0) * rotz(pi/2))

    else:
        RDK.setParam('prox_obj','NULL')

--- Python program Avanzar_Cinta_Rot ---
from robodk import *      # RoboDK API
from robolink import *    # Robot toolbox

RDK = Robolink()

cinta_rot=RDK.Item('Cinta_Rotativa',itemtype=ITEM_TYPE_ROBOT)

if cinta_rot.Valid():
    cinta_rot.MoveJ(cinta_rot.Joints()+220)
